(* IEC 61131-3 sources: trust-platform/examples/control/09-industrial-control-structures/60-loop-diagnosis/src, 1 file *)

(* ---- Main.st ---- *)
USING Control;

PROGRAM Main
VAR
    Controller : Control.PID;
    Parameters : Control.PIDParameters := (
        ProportionalGain := LREAL#2.0,
        IntegralGain := LREAL#0.5,
        DerivativeGain := LREAL#0.0,
        ProportionalSetpointWeight := LREAL#1.0,
        DerivativeSetpointWeight := LREAL#0.0,
        Bias := LREAL#0.0,
        OutputMinimum := LREAL#0.0,
        OutputMaximum := LREAL#100.0,
        RateMinimum := LREAL#-10000.0,
        RateMaximum := LREAL#10000.0,
        TrackingTime := LREAL#1.0,
        AntiWindup := PIDAntiWindup#BackCalculation
    );
    InitialState : Control.PIDInitialState;
    BeforeState : Control.PIDInitialState;
    ObservedState : Control.PIDInitialState;
    Input : Control.PIDInput;
    Initialized : BOOL := FALSE;
    ExperimentEnabled : BOOL := FALSE;
    HasStarted : BOOL := FALSE;
    SafetyAbort : BOOL := FALSE;
    AutoMode : BOOL := FALSE;
    TrialKind : INT := 0; (* 0:35→38°C target; 1:30kW extraction at SP35. *)
    KpPctPerC : LREAL := 2.0;
    KiPctPerCs : LREAL := 0.5;
    WaterTemperatureC : LREAL := 35.0;
    TemperatureC : LREAL := 35.0;
    SetpointC : LREAL := 35.0;
    DisturbanceKw : LREAL := 0.0;
    ErrorC : LREAL := 0.0;
    ProportionalPct : LREAL := 0.0;
    IntegralPct : LREAL := 75.0;
    RequestedPowerPct : LREAL := 75.0;
    HeaterCommandPct : LREAL := 75.0;
    AppliedPowerPct : LREAL := 75.0;
    PreviousRequestedPowerPct : LREAL := 75.0;
    PairedRequestPct : LREAL := 75.0;
    DiagnosticErrorC : LREAL := 0.0;
    ReferenceDifferenceC : LREAL := 0.0;
    UnavailableCommandPct : LREAL := 0.0;
    PositiveError : BOOL := FALSE;
    AtUpperLimit : BOOL := FALSE;
    ReferenceDisagrees : BOOL := FALSE;
END_VAR

(* One native process publishes measured temperature and an unbiased simulation
   reference through separate normal inputs. No plant or sensor effect is built here. *)
PairedRequestPct := PreviousRequestedPowerPct;
UnavailableCommandPct := PairedRequestPct - AppliedPowerPct;
IF NOT (TemperatureC >= LREAL#0.0 AND TemperatureC <= LREAL#80.0) THEN
    SafetyAbort := TRUE;
ELSE Input.ProcessValue := TemperatureC;
END_IF;
KpPctPerC := Parameters.ProportionalGain;
KiPctPerCs := Parameters.IntegralGain;
AutoMode := ExperimentEnabled AND NOT SafetyAbort;
SetpointC := LREAL#35.0;
DisturbanceKw := LREAL#0.0;
IF AutoMode THEN
    HasStarted := TRUE;
    IF TrialKind = 0 THEN SetpointC := LREAL#38.0;
    ELSIF TrialKind = 1 THEN DisturbanceKw := LREAL#30.0;
    END_IF;
    Input.Mode := PIDMode#Auto;
ELSE
    Input.Mode := PIDMode#Manual;
END_IF;
Input.ManualOutput := LREAL#0.0;
IF NOT HasStarted AND NOT SafetyAbort THEN Input.ManualOutput := LREAL#75.0;
END_IF;
Input.Setpoint := SetpointC;
Input.CycleTime := LREAL#0.1;
Input.FeedForward := LREAL#0.0;
Input.TrackingOutput := LREAL#0.0;
ErrorC := SetpointC - Input.ProcessValue;

Controller.Configure(Parameters := Parameters);
IF NOT Initialized THEN
    InitialState.Setpoint := LREAL#35.0;
    InitialState.ProcessValue := Input.ProcessValue;
    InitialState.NominalOutput := LREAL#75.0;
    InitialState.SaturatedOutput := LREAL#75.0;
    Controller.Initialize(State := InitialState);
    Initialized := TRUE;
END_IF;
BeforeState := Controller.GetState();

(* Fixed PI gains and weight one make nominal output = P + equivalent I.
   These observations use the library's retained state and own no actuator. *)
ProportionalPct := LREAL#0.0;
RequestedPowerPct := Input.ManualOutput;
IF AutoMode THEN
    ProportionalPct := KpPctPerC * ErrorC;
    RequestedPowerPct := BeforeState.NominalOutput
        + KpPctPerC * ((SetpointC - BeforeState.Setpoint)
            - (Input.ProcessValue - BeforeState.ProcessValue))
        + KiPctPerCs * ErrorC * Input.CycleTime;
END_IF;
HeaterCommandPct := Controller.Update(Input := Input);
ObservedState := Controller.GetState();
IntegralPct := ObservedState.NominalOutput - ProportionalPct;
PreviousRequestedPowerPct := RequestedPowerPct;

DiagnosticErrorC := SetpointC - TemperatureC;
ReferenceDifferenceC := TemperatureC - WaterTemperatureC;
PositiveError := DiagnosticErrorC > LREAL#0.0;
AtUpperLimit := AppliedPowerPct >= LREAL#100.0;
ReferenceDisagrees := ABS(ReferenceDifferenceC) > LREAL#0.2;
(* These remain separate observations, not an automatic capacity diagnosis.
   PairedRequestPct is the preceding request corresponding to this input scan;
   sensor acquisition timestamps and measured delivered kW remain unavailable. *)
END_PROGRAM

CONFIGURATION Config
RESOURCE Res ON PLC
    TASK MainTask(INTERVAL := T#100ms, PRIORITY := 1);
    PROGRAM P1 WITH MainTask : Main;
END_RESOURCE
VAR_CONFIG
    P1.ExperimentEnabled AT %MX112.0 : BOOL;
    P1.AutoMode AT %MX112.1 : BOOL;
    P1.SafetyAbort AT %MX112.2 : BOOL;
    P1.SetpointC AT %ML0 : LREAL;
    P1.ErrorC AT %ML8 : LREAL;
    P1.IntegralPct AT %ML16 : LREAL;
    P1.RequestedPowerPct AT %ML32 : LREAL;
    P1.WaterTemperatureC AT %IL16 : LREAL;
    P1.DiagnosticErrorC AT %ML64 : LREAL;
    P1.ReferenceDifferenceC AT %ML72 : LREAL;
    P1.UnavailableCommandPct AT %ML88 : LREAL;
    P1.PairedRequestPct AT %ML96 : LREAL;
    P1.PositiveError AT %MX120.0 : BOOL;
    P1.AtUpperLimit AT %MX120.1 : BOOL;
    P1.ReferenceDisagrees AT %MX120.2 : BOOL;
    P1.ProportionalPct AT %ML56 : LREAL;
    P1.TemperatureC AT %IL0 : LREAL;
    P1.AppliedPowerPct AT %IL8 : LREAL;
    P1.HeaterCommandPct AT %QL0 : LREAL;
    P1.DisturbanceKw AT %QL8 : LREAL;
END_VAR
END_CONFIGURATION
